(*
SPDX-FileCopyrightText: © 2026 Oleksandr Tiutyk <trofimich@gmail.com>
SPDX-License-Identifier: MIT
License: https://opensource.org/license/mit
*)

(*!
<summary>
Defines the contract for an activity that waits until an arbitrary workflow condition evaluates to TRUE.
</summary>
<description>
Advances cyclic execution until the associated condition evaluates to TRUE, then transitions to
PASSIVE_COMPLETED. Accepts simple, variable-based, composite (AND/OR), or custom condition implementations.
</description>
*)

INTERFACE IWaitConditionActivity EXTENDS IActivity

(*!
<summary>Returns the condition being evaluated, or 0 before configuration.</summary>
*)
{attribute 'monitoring' := 'call'}
PROPERTY Condition : ICondition
GET
END_GET
END_PROPERTY

(*!
<summary>Reports whether the condition has been configured.</summary>
*)
{attribute 'monitoring' := 'call'}
PROPERTY Configured : BOOL
GET
END_GET
END_PROPERTY

(*!
<summary>Configures the condition to wait for.</summary>
<description>
Validates that the condition is live, unattached to another parent, and establishes the parent link.
</description>
<param name="condition">Condition to evaluate during execution.</param>
*)
METHOD Configure
VAR_INPUT
	condition : ICondition;
END_VAR
END_METHOD

END_INTERFACE

(* stored: Version 1.1.0.1
   Itf IWaitConditionActivity: Id {0cefaf0d-4ae9-47b9-8f8d-e636a560d87a}
   Property Condition: Id {960bfa25-ba1a-4222-80a3-1359b946b290}
   Get Get: Id {4a9d6524-357e-4744-aaba-474fc163ec8b}
   Property Configured: Id {0ace7a5a-e627-4c38-8a84-290f9229d0de}
   Get Get: Id {db3ddcb3-657c-4070-be26-7ddb756d1f28}
   Method Configure: Id {142fa54f-1e2c-4c26-afda-45aa5107564f} *)
